TYPE ST_Banner_TL503Pro_Raw :
STRUCT
	PDOs	:	Array[20..30] of USINT;
END_STRUCT
END_TYPE

(* stored: Version 1.1.0.1
   DUT ST_Banner_TL503Pro_Raw: Id {b58958f7-bb51-4639-9bcc-c6f8a77e8315} *)
